(* IEC 61131-3 sources: sis-interlock-demo/tests/POUs/Generated/FB_CemGen02_Test, 41 files *)

(* ---- FB_CemGen02_Test.decl.st ---- *)
// AUTO-GENERATED by cemgen 1.0.0 — не редактировать: правьте матрицу и запустите
//   python -m cemgen generate <файл матрицы .csv или .xlsx>
// Матрица: SIS-V101-CEM, объект V-101, ревизия B от 2026-10-19, SHA-256 сетки df2ed4841a9453ca
// Назначение: набор coUnit: сценарии по матрице SIS-V101-CEM, тесты 41–80 (DESIGN.md, 12.4).
//             Ожидаемые значения — эталонная модель cemgen. Стенд FB_SisHarness — по экземпляру на
//             тест.
// Автор:      kr0nsch; код — генератор cemgen
// Версия:     1.0.0
// Документ:   docs/DESIGN.md, раздел «10. Генератор cemgen»; docs/cause_effect_matrix.md
// ВНИМАНИЕ:   код демонстрационный и не предназначен для систем безопасности. Реальная ПАЗ требует
//             определения SIL, сертифицированных аппаратных и программных средств и валидации по
//             ГОСТ Р МЭК 61511.
FUNCTION_BLOCK FB_CemGen02_Test EXTENDS coUnit.FB_TestSuite
VAR
    fbH001 : FB_SisHarness;   // Matrix_ASHH104Override_Denied
    fbH002 : FB_SisHarness;   // Matrix_ASHH104Reset_OnlyAfterClear
    fbH003 : FB_SisHarness;   // Matrix_ASHH104ChannelInvalid_MatchesPolicy
    fbH004 : FB_SisHarness;   // Matrix_ASHH104Bypass_ExpiresBackToVoting
    fbH005 : FB_SisHarness;   // Matrix_BSH105Demand_TripsOwnEffects
    fbH006 : FB_SisHarness;   // Matrix_BSH105Override_Denied
    fbH007 : FB_SisHarness;   // Matrix_BSH105Reset_OnlyAfterClear
    fbH008 : FB_SisHarness;   // Matrix_BSH105ChannelInvalid_MatchesPolicy
    fbH009 : FB_SisHarness;   // Matrix_BSH105Bypass_ExpiresBackToVoting
    fbH010 : FB_SisHarness;   // Matrix_HS106Demand_TripsOwnEffects
    fbH011 : FB_SisHarness;   // Matrix_HS106Override_Denied
    fbH012 : FB_SisHarness;   // Matrix_HS106Reset_OnlyAfterClear
    fbH013 : FB_SisHarness;   // Matrix_HS106ChannelInvalid_MatchesPolicy
    fbH014 : FB_SisHarness;   // Matrix_HS106Bypass_Denied
    fbH015 : FB_SisHarness;   // Matrix_PSLL108Demand_TripsOwnEffects
    fbH016 : FB_SisHarness;   // Matrix_PSLL108Delay_TripsExactlyAtDelay
    fbH017 : FB_SisHarness;   // Matrix_PSLL108Override_ExpiresThenTrips
    fbH018 : FB_SisHarness;   // Matrix_PSLL108Override_ClearsAfterConfirm
    fbH019 : FB_SisHarness;   // Matrix_PSLL108Override_DemandBackRestartsConfirm
    fbH020 : FB_SisHarness;   // Matrix_PSLL108Override_ExpiryBoundsConfirm
    fbH021 : FB_SisHarness;   // Matrix_PSLL108Override_ClearedThenDelayTrips
    fbH022 : FB_SisHarness;   // Matrix_PSLL108Reset_OnlyAfterClear
    fbH023 : FB_SisHarness;   // Matrix_PSLL108ChannelInvalid_MatchesPolicy
    fbH024 : FB_SisHarness;   // Matrix_PSLL108Bypass_ExpiresBackToVoting
    fbH025 : FB_SisHarness;   // Matrix_ESL109Demand_TripsOwnEffects
    fbH026 : FB_SisHarness;   // Matrix_ESL109Delay_TripsExactlyAtDelay
    fbH027 : FB_SisHarness;   // Matrix_ESL109Override_Denied
    fbH028 : FB_SisHarness;   // Matrix_ESL109Reset_OnlyAfterClear
    fbH029 : FB_SisHarness;   // Matrix_ESL109ChannelInvalid_MatchesPolicy
    fbH030 : FB_SisHarness;   // Matrix_ESL109Bypass_Denied
    fbH031 : FB_SisHarness;   // Matrix_FirstOutPSHH101ThenPSLL101_RecordsFirst
    fbH032 : FB_SisHarness;   // Matrix_FirstOutPSLL101ThenLSHH102_RecordsFirst
    fbH033 : FB_SisHarness;   // Matrix_FirstOutLSHH102ThenLSLL102_RecordsFirst
    fbH034 : FB_SisHarness;   // Matrix_FirstOutLSLL102ThenTSHH103_RecordsFirst
    fbH035 : FB_SisHarness;   // Matrix_FirstOutTSHH103ThenASHH104_RecordsFirst
    fbH036 : FB_SisHarness;   // Matrix_FirstOutASHH104ThenBSH105_RecordsFirst
    fbH037 : FB_SisHarness;   // Matrix_FirstOutBSH105ThenHS106_RecordsFirst
    fbH038 : FB_SisHarness;   // Matrix_FirstOutHS106ThenPSLL108_RecordsFirst
    fbH039 : FB_SisHarness;   // Matrix_FirstOutPSLL108ThenESL109_RecordsFirst
    fbH040 : FB_SisHarness;   // Matrix_FirstOutESL109ThenPSHH101_RecordsFirst
END_VAR

(* ---- ASHH104BypassExpiresBackToVoting.method.decl.st ---- *)
// AUTO-GENERATED by cemgen 1.0.0 — не редактировать: правьте матрицу и запустите
//   python -m cemgen generate <файл матрицы .csv или .xlsx>
// Матрица: SIS-V101-CEM, объект V-101, ревизия B от 2026-10-19, SHA-256 сетки df2ed4841a9453ca
// Назначение: тест Matrix_ASHH104Bypass_ExpiresBackToVoting набора FB_CemGen02_Test (сценарий по
//             матрице, DESIGN.md, 12.4).
// Автор:      kr0nsch; код — генератор cemgen
// Версия:     1.0.0
// Документ:   docs/DESIGN.md, раздел «10. Генератор cemgen»; docs/cause_effect_matrix.md
// ВНИМАНИЕ:   код демонстрационный и не предназначен для систем безопасности. Реальная ПАЗ требует
//             определения SIL, сертифицированных аппаратных и программных средств и валидации по
//             ГОСТ Р МЭК 61511.
// Причина 6 ASHH104: ключ разрешения байпасов, байпас AT104A → Active; канал недостоверен → Bypassed,
// не сработало; на t0 + 8 ч − шаг — Active; ровно на t0 + 8 ч — Expired, BypassExpired, канал Invalid;
// далее — по эталонной модели.
METHOD PRIVATE ASHH104BypassExpiresBackToVoting
VAR
    xArmed : BOOL;           // стенд взведён: все следствия под напряжением после сброса
    stVs   : ST_VotingSts;   // копия состояния группы голосования
END_VAR

(* ---- ASHH104ChannelInvalidMatchesPolicy.method.decl.st ---- *)
// AUTO-GENERATED by cemgen 1.0.0 — не редактировать: правьте матрицу и запустите
//   python -m cemgen generate <файл матрицы .csv или .xlsx>
// Матрица: SIS-V101-CEM, объект V-101, ревизия B от 2026-10-19, SHA-256 сетки df2ed4841a9453ca
// Назначение: тест Matrix_ASHH104ChannelInvalid_MatchesPolicy набора FB_CemGen02_Test (сценарий по
//             матрице, DESIGN.md, 12.4).
// Автор:      kr0nsch; код — генератор cemgen
// Версия:     1.0.0
// Документ:   docs/DESIGN.md, раздел «10. Генератор cemgen»; docs/cause_effect_matrix.md
// ВНИМАНИЕ:   код демонстрационный и не предназначен для систем безопасности. Реальная ПАЗ требует
//             определения SIL, сертифицированных аппаратных и программных средств и валидации по
//             ГОСТ Р МЭК 61511.
// Причина 6 ASHH104 (2oo3, DegradeSafe): канал AT104A недостоверен → действующая схема и срабатывание
// по политике деградации; если не сработало — требование на AT104B → по эталонной модели.
METHOD PRIVATE ASHH104ChannelInvalidMatchesPolicy
VAR
    xArmed : BOOL;           // стенд взведён: все следствия под напряжением после сброса
    stVs   : ST_VotingSts;   // копия состояния группы голосования
END_VAR

(* ---- ASHH104OverrideDenied.method.decl.st ---- *)
// AUTO-GENERATED by cemgen 1.0.0 — не редактировать: правьте матрицу и запустите
//   python -m cemgen generate <файл матрицы .csv или .xlsx>
// Матрица: SIS-V101-CEM, объект V-101, ревизия B от 2026-10-19, SHA-256 сетки df2ed4841a9453ca
// Назначение: тест Matrix_ASHH104Override_Denied набора FB_CemGen02_Test (сценарий по матрице,
//             DESIGN.md, 12.4).
// Автор:      kr0nsch; код — генератор cemgen
// Версия:     1.0.0
// Документ:   docs/DESIGN.md, раздел «10. Генератор cemgen»; docs/cause_effect_matrix.md
// ВНИМАНИЕ:   код демонстрационный и не предназначен для систем безопасности. Реальная ПАЗ требует
//             определения SIL, сертифицированных аппаратных и программных средств и валидации по
//             ГОСТ Р МЭК 61511.
// Причина 6 ASHH104 без разрешённого обхода: ключ разрешения обходов, запрос → последнее событие
// OverrideDenied, обхода нет; требование → срабатывание после задержки.
METHOD PRIVATE ASHH104OverrideDenied
VAR
    xArmed : BOOL;          // стенд взведён: все следствия под напряжением после сброса
    stEv   : ST_SisEvent;   // последнее событие журнала
END_VAR

(* ---- ASHH104ResetOnlyAfterClear.method.decl.st ---- *)
// AUTO-GENERATED by cemgen 1.0.0 — не редактировать: правьте матрицу и запустите
//   python -m cemgen generate <файл матрицы .csv или .xlsx>
// Матрица: SIS-V101-CEM, объект V-101, ревизия B от 2026-10-19, SHA-256 сетки df2ed4841a9453ca
// Назначение: тест Matrix_ASHH104Reset_OnlyAfterClear набора FB_CemGen02_Test (сценарий по матрице,
//             DESIGN.md, 12.4).
// Автор:      kr0nsch; код — генератор cemgen
// Версия:     1.0.0
// Документ:   docs/DESIGN.md, раздел «10. Генератор cemgen»; docs/cause_effect_matrix.md
// ВНИМАНИЕ:   код демонстрационный и не предназначен для систем безопасности. Реальная ПАЗ требует
//             определения SIL, сертифицированных аппаратных и программных средств и валидации по
//             ГОСТ Р МЭК 61511.
// Причина 6 ASHH104: срабатывание; сброс при требовании → ResetDenied, блокирует ASHH104, следствия
// обесточены; норма → следствия всё ещё обесточены (фиксация); сброс → все следствия под напряжением.
METHOD PRIVATE ASHH104ResetOnlyAfterClear
VAR
    xArmed : BOOL;          // стенд взведён: все следствия под напряжением после сброса
    stEv   : ST_SisEvent;   // последнее событие журнала
END_VAR

(* ---- BSH105BypassExpiresBackToVoting.method.decl.st ---- *)
// AUTO-GENERATED by cemgen 1.0.0 — не редактировать: правьте матрицу и запустите
//   python -m cemgen generate <файл матрицы .csv или .xlsx>
// Матрица: SIS-V101-CEM, объект V-101, ревизия B от 2026-10-19, SHA-256 сетки df2ed4841a9453ca
// Назначение: тест Matrix_BSH105Bypass_ExpiresBackToVoting набора FB_CemGen02_Test (сценарий по
//             матрице, DESIGN.md, 12.4).
// Автор:      kr0nsch; код — генератор cemgen
// Версия:     1.0.0
// Документ:   docs/DESIGN.md, раздел «10. Генератор cemgen»; docs/cause_effect_matrix.md
// ВНИМАНИЕ:   код демонстрационный и не предназначен для систем безопасности. Реальная ПАЗ требует
//             определения SIL, сертифицированных аппаратных и программных средств и валидации по
//             ГОСТ Р МЭК 61511.
// Причина 7 BSH105: ключ разрешения байпасов, байпас BS105A → Active; канал недостоверен → Bypassed,
// не сработало; на t0 + 8 ч − шаг — Active; ровно на t0 + 8 ч — Expired, BypassExpired, канал Invalid;
// далее — по эталонной модели.
METHOD PRIVATE BSH105BypassExpiresBackToVoting
VAR
    xArmed : BOOL;           // стенд взведён: все следствия под напряжением после сброса
    stVs   : ST_VotingSts;   // копия состояния группы голосования
END_VAR

(* ---- BSH105ChannelInvalidMatchesPolicy.method.decl.st ---- *)
// AUTO-GENERATED by cemgen 1.0.0 — не редактировать: правьте матрицу и запустите
//   python -m cemgen generate <файл матрицы .csv или .xlsx>
// Матрица: SIS-V101-CEM, объект V-101, ревизия B от 2026-10-19, SHA-256 сетки df2ed4841a9453ca
// Назначение: тест Matrix_BSH105ChannelInvalid_MatchesPolicy набора FB_CemGen02_Test (сценарий по
//             матрице, DESIGN.md, 12.4).
// Автор:      kr0nsch; код — генератор cemgen
// Версия:     1.0.0
// Документ:   docs/DESIGN.md, раздел «10. Генератор cemgen»; docs/cause_effect_matrix.md
// ВНИМАНИЕ:   код демонстрационный и не предназначен для систем безопасности. Реальная ПАЗ требует
//             определения SIL, сертифицированных аппаратных и программных средств и валидации по
//             ГОСТ Р МЭК 61511.
// Причина 7 BSH105 (1oo2, DegradeSafe): канал BS105A недостоверен → действующая схема и срабатывание
// по политике деградации; если не сработало — требование на BS105B → по эталонной модели.
METHOD PRIVATE BSH105ChannelInvalidMatchesPolicy
VAR
    xArmed : BOOL;           // стенд взведён: все следствия под напряжением после сброса
    stVs   : ST_VotingSts;   // копия состояния группы голосования
END_VAR

(* ---- BSH105DemandTripsOwnEffects.method.decl.st ---- *)
// AUTO-GENERATED by cemgen 1.0.0 — не редактировать: правьте матрицу и запустите
//   python -m cemgen generate <файл матрицы .csv или .xlsx>
// Матрица: SIS-V101-CEM, объект V-101, ревизия B от 2026-10-19, SHA-256 сетки df2ed4841a9453ca
// Назначение: тест Matrix_BSH105Demand_TripsOwnEffects набора FB_CemGen02_Test (сценарий по
//             матрице, DESIGN.md, 12.4).
// Автор:      kr0nsch; код — генератор cemgen
// Версия:     1.0.0
// Документ:   docs/DESIGN.md, раздел «10. Генератор cemgen»; docs/cause_effect_matrix.md
// ВНИМАНИЕ:   код демонстрационный и не предназначен для систем безопасности. Реальная ПАЗ требует
//             определения SIL, сертифицированных аппаратных и программных средств и валидации по
//             ГОСТ Р МЭК 61511.
// Причина 7 BSH105 (1oo2, задержка 0 с): требование BS105A, BS105B = 0 отключает ESDV101, BDV101,
// ESDV102, P101A, P101B, H101, UA110; остальные следствия под напряжением; первопричина BSH105.
METHOD PRIVATE BSH105DemandTripsOwnEffects
VAR
    xArmed : BOOL;   // стенд взведён: все следствия под напряжением после сброса
END_VAR

(* ---- BSH105OverrideDenied.method.decl.st ---- *)
// AUTO-GENERATED by cemgen 1.0.0 — не редактировать: правьте матрицу и запустите
//   python -m cemgen generate <файл матрицы .csv или .xlsx>
// Матрица: SIS-V101-CEM, объект V-101, ревизия B от 2026-10-19, SHA-256 сетки df2ed4841a9453ca
// Назначение: тест Matrix_BSH105Override_Denied набора FB_CemGen02_Test (сценарий по матрице,
//             DESIGN.md, 12.4).
// Автор:      kr0nsch; код — генератор cemgen
// Версия:     1.0.0
// Документ:   docs/DESIGN.md, раздел «10. Генератор cemgen»; docs/cause_effect_matrix.md
// ВНИМАНИЕ:   код демонстрационный и не предназначен для систем безопасности. Реальная ПАЗ требует
//             определения SIL, сертифицированных аппаратных и программных средств и валидации по
//             ГОСТ Р МЭК 61511.
// Причина 7 BSH105 без разрешённого обхода: ключ разрешения обходов, запрос → последнее событие
// OverrideDenied, обхода нет; требование → срабатывание после задержки.
METHOD PRIVATE BSH105OverrideDenied
VAR
    xArmed : BOOL;          // стенд взведён: все следствия под напряжением после сброса
    stEv   : ST_SisEvent;   // последнее событие журнала
END_VAR

(* ---- BSH105ResetOnlyAfterClear.method.decl.st ---- *)
// AUTO-GENERATED by cemgen 1.0.0 — не редактировать: правьте матрицу и запустите
//   python -m cemgen generate <файл матрицы .csv или .xlsx>
// Матрица: SIS-V101-CEM, объект V-101, ревизия B от 2026-10-19, SHA-256 сетки df2ed4841a9453ca
// Назначение: тест Matrix_BSH105Reset_OnlyAfterClear набора FB_CemGen02_Test (сценарий по матрице,
//             DESIGN.md, 12.4).
// Автор:      kr0nsch; код — генератор cemgen
// Версия:     1.0.0
// Документ:   docs/DESIGN.md, раздел «10. Генератор cemgen»; docs/cause_effect_matrix.md
// ВНИМАНИЕ:   код демонстрационный и не предназначен для систем безопасности. Реальная ПАЗ требует
//             определения SIL, сертифицированных аппаратных и программных средств и валидации по
//             ГОСТ Р МЭК 61511.
// Причина 7 BSH105: срабатывание; сброс при требовании → ResetDenied, блокирует BSH105, следствия
// обесточены; норма → следствия всё ещё обесточены (фиксация); сброс → все следствия под напряжением.
METHOD PRIVATE BSH105ResetOnlyAfterClear
VAR
    xArmed : BOOL;          // стенд взведён: все следствия под напряжением после сброса
    stEv   : ST_SisEvent;   // последнее событие журнала
END_VAR

(* ---- ESL109BypassDenied.method.decl.st ---- *)
// AUTO-GENERATED by cemgen 1.0.0 — не редактировать: правьте матрицу и запустите
//   python -m cemgen generate <файл матрицы .csv или .xlsx>
// Матрица: SIS-V101-CEM, объект V-101, ревизия B от 2026-10-19, SHA-256 сетки df2ed4841a9453ca
// Назначение: тест Matrix_ESL109Bypass_Denied набора FB_CemGen02_Test (сценарий по матрице,
//             DESIGN.md, 12.4).
// Автор:      kr0nsch; код — генератор cemgen
// Версия:     1.0.0
// Документ:   docs/DESIGN.md, раздел «10. Генератор cemgen»; docs/cause_effect_matrix.md
// ВНИМАНИЕ:   код демонстрационный и не предназначен для систем безопасности. Реальная ПАЗ требует
//             определения SIL, сертифицированных аппаратных и программных средств и валидации по
//             ГОСТ Р МЭК 61511.
// Причина 10 ESL109: байпас запрещён (bypass_max = 0); ключ разрешения байпасов, запрос байпаса ES109
// → Denied, событие BypassDenied с номером канала.
METHOD PRIVATE ESL109BypassDenied
VAR
    xArmed : BOOL;           // стенд взведён: все следствия под напряжением после сброса
    stVs   : ST_VotingSts;   // копия состояния группы голосования
    stEv   : ST_SisEvent;    // последнее событие журнала
END_VAR

(* ---- ESL109ChannelInvalidMatchesPolicy.method.decl.st ---- *)
// AUTO-GENERATED by cemgen 1.0.0 — не редактировать: правьте матрицу и запустите
//   python -m cemgen generate <файл матрицы .csv или .xlsx>
// Матрица: SIS-V101-CEM, объект V-101, ревизия B от 2026-10-19, SHA-256 сетки df2ed4841a9453ca
// Назначение: тест Matrix_ESL109ChannelInvalid_MatchesPolicy набора FB_CemGen02_Test (сценарий по
//             матрице, DESIGN.md, 12.4).
// Автор:      kr0nsch; код — генератор cemgen
// Версия:     1.0.0
// Документ:   docs/DESIGN.md, раздел «10. Генератор cemgen»; docs/cause_effect_matrix.md
// ВНИМАНИЕ:   код демонстрационный и не предназначен для систем безопасности. Реальная ПАЗ требует
//             определения SIL, сертифицированных аппаратных и программных средств и валидации по
//             ГОСТ Р МЭК 61511.
// Причина 10 ESL109 (1oo1, VoteTrip): канал ES109 недостоверен → действующая схема и срабатывание по
// политике деградации; если не сработало — требование на втором канале → по эталонной модели.
METHOD PRIVATE ESL109ChannelInvalidMatchesPolicy
VAR
    xArmed : BOOL;           // стенд взведён: все следствия под напряжением после сброса
    stVs   : ST_VotingSts;   // копия состояния группы голосования
END_VAR

(* ---- ESL109DelayTripsExactlyAtDelay.method.decl.st ---- *)
// AUTO-GENERATED by cemgen 1.0.0 — не редактировать: правьте матрицу и запустите
//   python -m cemgen generate <файл матрицы .csv или .xlsx>
// Матрица: SIS-V101-CEM, объект V-101, ревизия B от 2026-10-19, SHA-256 сетки df2ed4841a9453ca
// Назначение: тест Matrix_ESL109Delay_TripsExactlyAtDelay набора FB_CemGen02_Test (сценарий по
//             матрице, DESIGN.md, 12.4).
// Автор:      kr0nsch; код — генератор cemgen
// Версия:     1.0.0
// Документ:   docs/DESIGN.md, раздел «10. Генератор cemgen»; docs/cause_effect_matrix.md
// ВНИМАНИЕ:   код демонстрационный и не предназначен для систем безопасности. Реальная ПАЗ требует
//             определения SIL, сертифицированных аппаратных и программных средств и валидации по
//             ГОСТ Р МЭК 61511.
// Причина 10 ESL109: требование в t0; на t0 + 2 с − шаг не зафиксирована, следствия под напряжением;
// ровно на t0 + 2 с — зафиксирована, ltFirstOut = t0 + задержка.
METHOD PRIVATE ESL109DelayTripsExactlyAtDelay
VAR
    xArmed : BOOL;    // стенд взведён: все следствия под напряжением после сброса
    ltT0   : LTIME;   // момент t0 по подменному времени стенда
END_VAR

(* ---- ESL109DemandTripsOwnEffects.method.decl.st ---- *)
// AUTO-GENERATED by cemgen 1.0.0 — не редактировать: правьте матрицу и запустите
//   python -m cemgen generate <файл матрицы .csv или .xlsx>
// Матрица: SIS-V101-CEM, объект V-101, ревизия B от 2026-10-19, SHA-256 сетки df2ed4841a9453ca
// Назначение: тест Matrix_ESL109Demand_TripsOwnEffects набора FB_CemGen02_Test (сценарий по
//             матрице, DESIGN.md, 12.4).
// Автор:      kr0nsch; код — генератор cemgen
// Версия:     1.0.0
// Документ:   docs/DESIGN.md, раздел «10. Генератор cemgen»; docs/cause_effect_matrix.md
// ВНИМАНИЕ:   код демонстрационный и не предназначен для систем безопасности. Реальная ПАЗ требует
//             определения SIL, сертифицированных аппаратных и программных средств и валидации по
//             ГОСТ Р МЭК 61511.
// Причина 10 ESL109 (1oo1, задержка 2 с): требование ES109 = 0 отключает P101A, P101B, H101, UA110;
// остальные следствия под напряжением; первопричина ESL109.
METHOD PRIVATE ESL109DemandTripsOwnEffects
VAR
    xArmed : BOOL;   // стенд взведён: все следствия под напряжением после сброса
END_VAR

(* ---- ESL109OverrideDenied.method.decl.st ---- *)
// AUTO-GENERATED by cemgen 1.0.0 — не редактировать: правьте матрицу и запустите
//   python -m cemgen generate <файл матрицы .csv или .xlsx>
// Матрица: SIS-V101-CEM, объект V-101, ревизия B от 2026-10-19, SHA-256 сетки df2ed4841a9453ca
// Назначение: тест Matrix_ESL109Override_Denied набора FB_CemGen02_Test (сценарий по матрице,
//             DESIGN.md, 12.4).
// Автор:      kr0nsch; код — генератор cemgen
// Версия:     1.0.0
// Документ:   docs/DESIGN.md, раздел «10. Генератор cemgen»; docs/cause_effect_matrix.md
// ВНИМАНИЕ:   код демонстрационный и не предназначен для систем безопасности. Реальная ПАЗ требует
//             определения SIL, сертифицированных аппаратных и программных средств и валидации по
//             ГОСТ Р МЭК 61511.
// Причина 10 ESL109 без разрешённого обхода: ключ разрешения обходов, запрос → последнее событие
// OverrideDenied, обхода нет; требование → срабатывание после задержки.
METHOD PRIVATE ESL109OverrideDenied
VAR
    xArmed : BOOL;          // стенд взведён: все следствия под напряжением после сброса
    stEv   : ST_SisEvent;   // последнее событие журнала
END_VAR

(* ---- ESL109ResetOnlyAfterClear.method.decl.st ---- *)
// AUTO-GENERATED by cemgen 1.0.0 — не редактировать: правьте матрицу и запустите
//   python -m cemgen generate <файл матрицы .csv или .xlsx>
// Матрица: SIS-V101-CEM, объект V-101, ревизия B от 2026-10-19, SHA-256 сетки df2ed4841a9453ca
// Назначение: тест Matrix_ESL109Reset_OnlyAfterClear набора FB_CemGen02_Test (сценарий по матрице,
//             DESIGN.md, 12.4).
// Автор:      kr0nsch; код — генератор cemgen
// Версия:     1.0.0
// Документ:   docs/DESIGN.md, раздел «10. Генератор cemgen»; docs/cause_effect_matrix.md
// ВНИМАНИЕ:   код демонстрационный и не предназначен для систем безопасности. Реальная ПАЗ требует
//             определения SIL, сертифицированных аппаратных и программных средств и валидации по
//             ГОСТ Р МЭК 61511.
// Причина 10 ESL109: срабатывание; сброс при требовании → ResetDenied, блокирует ESL109, следствия
// обесточены; норма → следствия всё ещё обесточены (фиксация); сброс → все следствия под напряжением.
METHOD PRIVATE ESL109ResetOnlyAfterClear
VAR
    xArmed : BOOL;          // стенд взведён: все следствия под напряжением после сброса
    stEv   : ST_SisEvent;   // последнее событие журнала
END_VAR

(* ---- FirstOutASHH104ThenBSH105RecordsFirst.method.decl.st ---- *)
// AUTO-GENERATED by cemgen 1.0.0 — не редактировать: правьте матрицу и запустите
//   python -m cemgen generate <файл матрицы .csv или .xlsx>
// Матрица: SIS-V101-CEM, объект V-101, ревизия B от 2026-10-19, SHA-256 сетки df2ed4841a9453ca
// Назначение: тест Matrix_FirstOutASHH104ThenBSH105_RecordsFirst набора FB_CemGen02_Test (сценарий
//             по матрице, DESIGN.md, 12.4).
// Автор:      kr0nsch; код — генератор cemgen
// Версия:     1.0.0
// Документ:   docs/DESIGN.md, раздел «10. Генератор cemgen»; docs/cause_effect_matrix.md
// ВНИМАНИЕ:   код демонстрационный и не предназначен для систем безопасности. Реальная ПАЗ требует
//             определения SIL, сертифицированных аппаратных и программных средств и валидации по
//             ГОСТ Р МЭК 61511.
// Первопричина: требование ASHH104, фиксация через 2 с; затем требование BSH105, фиксация через 0 с →
// первопричина ASHH104, в маске первопричины только ASHH104, ltFirstOut — момент фиксации ASHH104,
// BSH105 — среди зафиксированных.
METHOD PRIVATE FirstOutASHH104ThenBSH105RecordsFirst
VAR
    xArmed : BOOL;    // стенд взведён: все следствия под напряжением после сброса
    ltT0   : LTIME;   // момент t0 по подменному времени стенда
END_VAR

(* ---- FirstOutBSH105ThenHS106RecordsFirst.method.decl.st ---- *)
// AUTO-GENERATED by cemgen 1.0.0 — не редактировать: правьте матрицу и запустите
//   python -m cemgen generate <файл матрицы .csv или .xlsx>
// Матрица: SIS-V101-CEM, объект V-101, ревизия B от 2026-10-19, SHA-256 сетки df2ed4841a9453ca
// Назначение: тест Matrix_FirstOutBSH105ThenHS106_RecordsFirst набора FB_CemGen02_Test (сценарий по
//             матрице, DESIGN.md, 12.4).
// Автор:      kr0nsch; код — генератор cemgen
// Версия:     1.0.0
// Документ:   docs/DESIGN.md, раздел «10. Генератор cemgen»; docs/cause_effect_matrix.md
// ВНИМАНИЕ:   код демонстрационный и не предназначен для систем безопасности. Реальная ПАЗ требует
//             определения SIL, сертифицированных аппаратных и программных средств и валидации по
//             ГОСТ Р МЭК 61511.
// Первопричина: требование BSH105, фиксация через 0 с; затем требование HS106, фиксация через 0 с →
// первопричина BSH105, в маске первопричины только BSH105, ltFirstOut — момент фиксации BSH105, HS106
// — среди зафиксированных.
METHOD PRIVATE FirstOutBSH105ThenHS106RecordsFirst
VAR
    xArmed : BOOL;    // стенд взведён: все следствия под напряжением после сброса
    ltT0   : LTIME;   // момент t0 по подменному времени стенда
END_VAR

(* ---- FirstOutESL109ThenPSHH101RecordsFirst.method.decl.st ---- *)
// AUTO-GENERATED by cemgen 1.0.0 — не редактировать: правьте матрицу и запустите
//   python -m cemgen generate <файл матрицы .csv или .xlsx>
// Матрица: SIS-V101-CEM, объект V-101, ревизия B от 2026-10-19, SHA-256 сетки df2ed4841a9453ca
// Назначение: тест Matrix_FirstOutESL109ThenPSHH101_RecordsFirst набора FB_CemGen02_Test (сценарий
//             по матрице, DESIGN.md, 12.4).
// Автор:      kr0nsch; код — генератор cemgen
// Версия:     1.0.0
// Документ:   docs/DESIGN.md, раздел «10. Генератор cemgen»; docs/cause_effect_matrix.md
// ВНИМАНИЕ:   код демонстрационный и не предназначен для систем безопасности. Реальная ПАЗ требует
//             определения SIL, сертифицированных аппаратных и программных средств и валидации по
//             ГОСТ Р МЭК 61511.
// Первопричина: требование ESL109, фиксация через 2 с; затем требование PSHH101, фиксация через 2 с →
// первопричина ESL109, в маске первопричины только ESL109, ltFirstOut — момент фиксации ESL109,
// PSHH101 — среди зафиксированных.
METHOD PRIVATE FirstOutESL109ThenPSHH101RecordsFirst
VAR
    xArmed : BOOL;    // стенд взведён: все следствия под напряжением после сброса
    ltT0   : LTIME;   // момент t0 по подменному времени стенда
END_VAR

(* ---- FirstOutHS106ThenPSLL108RecordsFirst.method.decl.st ---- *)
// AUTO-GENERATED by cemgen 1.0.0 — не редактировать: правьте матрицу и запустите
//   python -m cemgen generate <файл матрицы .csv или .xlsx>
// Матрица: SIS-V101-CEM, объект V-101, ревизия B от 2026-10-19, SHA-256 сетки df2ed4841a9453ca
// Назначение: тест Matrix_FirstOutHS106ThenPSLL108_RecordsFirst набора FB_CemGen02_Test (сценарий
//             по матрице, DESIGN.md, 12.4).
// Автор:      kr0nsch; код — генератор cemgen
// Версия:     1.0.0
// Документ:   docs/DESIGN.md, раздел «10. Генератор cemgen»; docs/cause_effect_matrix.md
// ВНИМАНИЕ:   код демонстрационный и не предназначен для систем безопасности. Реальная ПАЗ требует
//             определения SIL, сертифицированных аппаратных и программных средств и валидации по
//             ГОСТ Р МЭК 61511.
// Первопричина: требование HS106, фиксация через 0 с; затем требование PSLL108, фиксация через 10 с →
// первопричина HS106, в маске первопричины только HS106, ltFirstOut — момент фиксации HS106, PSLL108 —
// среди зафиксированных.
METHOD PRIVATE FirstOutHS106ThenPSLL108RecordsFirst
VAR
    xArmed : BOOL;    // стенд взведён: все следствия под напряжением после сброса
    ltT0   : LTIME;   // момент t0 по подменному времени стенда
END_VAR

(* ---- FirstOutLSHH102ThenLSLL102RecordsFirst.method.decl.st ---- *)
// AUTO-GENERATED by cemgen 1.0.0 — не редактировать: правьте матрицу и запустите
//   python -m cemgen generate <файл матрицы .csv или .xlsx>
// Матрица: SIS-V101-CEM, объект V-101, ревизия B от 2026-10-19, SHA-256 сетки df2ed4841a9453ca
// Назначение: тест Matrix_FirstOutLSHH102ThenLSLL102_RecordsFirst набора FB_CemGen02_Test (сценарий
//             по матрице, DESIGN.md, 12.4).
// Автор:      kr0nsch; код — генератор cemgen
// Версия:     1.0.0
// Документ:   docs/DESIGN.md, раздел «10. Генератор cemgen»; docs/cause_effect_matrix.md
// ВНИМАНИЕ:   код демонстрационный и не предназначен для систем безопасности. Реальная ПАЗ требует
//             определения SIL, сертифицированных аппаратных и программных средств и валидации по
//             ГОСТ Р МЭК 61511.
// Первопричина: требование LSHH102, фиксация через 3 с; затем требование LSLL102, фиксация через 5 с →
// первопричина LSHH102, в маске первопричины только LSHH102, ltFirstOut — момент фиксации LSHH102,
// LSLL102 — среди зафиксированных.
METHOD PRIVATE FirstOutLSHH102ThenLSLL102RecordsFirst
VAR
    xArmed : BOOL;    // стенд взведён: все следствия под напряжением после сброса
    ltT0   : LTIME;   // момент t0 по подменному времени стенда
END_VAR

(* ---- FirstOutLSLL102ThenTSHH103RecordsFirst.method.decl.st ---- *)
// AUTO-GENERATED by cemgen 1.0.0 — не редактировать: правьте матрицу и запустите
//   python -m cemgen generate <файл матрицы .csv или .xlsx>
// Матрица: SIS-V101-CEM, объект V-101, ревизия B от 2026-10-19, SHA-256 сетки df2ed4841a9453ca
// Назначение: тест Matrix_FirstOutLSLL102ThenTSHH103_RecordsFirst набора FB_CemGen02_Test (сценарий
//             по матрице, DESIGN.md, 12.4).
// Автор:      kr0nsch; код — генератор cemgen
// Версия:     1.0.0
// Документ:   docs/DESIGN.md, раздел «10. Генератор cemgen»; docs/cause_effect_matrix.md
// ВНИМАНИЕ:   код демонстрационный и не предназначен для систем безопасности. Реальная ПАЗ требует
//             определения SIL, сертифицированных аппаратных и программных средств и валидации по
//             ГОСТ Р МЭК 61511.
// Первопричина: требование LSLL102, фиксация через 5 с; затем требование TSHH103, фиксация через 5 с →
// первопричина LSLL102, в маске первопричины только LSLL102, ltFirstOut — момент фиксации LSLL102,
// TSHH103 — среди зафиксированных.
METHOD PRIVATE FirstOutLSLL102ThenTSHH103RecordsFirst
VAR
    xArmed : BOOL;    // стенд взведён: все следствия под напряжением после сброса
    ltT0   : LTIME;   // момент t0 по подменному времени стенда
END_VAR

(* ---- FirstOutPSHH101ThenPSLL101RecordsFirst.method.decl.st ---- *)
// AUTO-GENERATED by cemgen 1.0.0 — не редактировать: правьте матрицу и запустите
//   python -m cemgen generate <файл матрицы .csv или .xlsx>
// Матрица: SIS-V101-CEM, объект V-101, ревизия B от 2026-10-19, SHA-256 сетки df2ed4841a9453ca
// Назначение: тест Matrix_FirstOutPSHH101ThenPSLL101_RecordsFirst набора FB_CemGen02_Test (сценарий
//             по матрице, DESIGN.md, 12.4).
// Автор:      kr0nsch; код — генератор cemgen
// Версия:     1.0.0
// Документ:   docs/DESIGN.md, раздел «10. Генератор cemgen»; docs/cause_effect_matrix.md
// ВНИМАНИЕ:   код демонстрационный и не предназначен для систем безопасности. Реальная ПАЗ требует
//             определения SIL, сертифицированных аппаратных и программных средств и валидации по
//             ГОСТ Р МЭК 61511.
// Первопричина: требование PSHH101, фиксация через 2 с; затем требование PSLL101, фиксация через 5 с →
// первопричина PSHH101, в маске первопричины только PSHH101, ltFirstOut — момент фиксации PSHH101,
// PSLL101 — среди зафиксированных.
METHOD PRIVATE FirstOutPSHH101ThenPSLL101RecordsFirst
VAR
    xArmed : BOOL;    // стенд взведён: все следствия под напряжением после сброса
    ltT0   : LTIME;   // момент t0 по подменному времени стенда
END_VAR

(* ---- FirstOutPSLL101ThenLSHH102RecordsFirst.method.decl.st ---- *)
// AUTO-GENERATED by cemgen 1.0.0 — не редактировать: правьте матрицу и запустите
//   python -m cemgen generate <файл матрицы .csv или .xlsx>
// Матрица: SIS-V101-CEM, объект V-101, ревизия B от 2026-10-19, SHA-256 сетки df2ed4841a9453ca
// Назначение: тест Matrix_FirstOutPSLL101ThenLSHH102_RecordsFirst набора FB_CemGen02_Test (сценарий
//             по матрице, DESIGN.md, 12.4).
// Автор:      kr0nsch; код — генератор cemgen
// Версия:     1.0.0
// Документ:   docs/DESIGN.md, раздел «10. Генератор cemgen»; docs/cause_effect_matrix.md
// ВНИМАНИЕ:   код демонстрационный и не предназначен для систем безопасности. Реальная ПАЗ требует
//             определения SIL, сертифицированных аппаратных и программных средств и валидации по
//             ГОСТ Р МЭК 61511.
// Первопричина: требование PSLL101, фиксация через 5 с; затем требование LSHH102, фиксация через 3 с →
// первопричина PSLL101, в маске первопричины только PSLL101, ltFirstOut — момент фиксации PSLL101,
// LSHH102 — среди зафиксированных.
METHOD PRIVATE FirstOutPSLL101ThenLSHH102RecordsFirst
VAR
    xArmed : BOOL;    // стенд взведён: все следствия под напряжением после сброса
    ltT0   : LTIME;   // момент t0 по подменному времени стенда
END_VAR

(* ---- FirstOutPSLL108ThenESL109RecordsFirst.method.decl.st ---- *)
// AUTO-GENERATED by cemgen 1.0.0 — не редактировать: правьте матрицу и запустите
//   python -m cemgen generate <файл матрицы .csv или .xlsx>
// Матрица: SIS-V101-CEM, объект V-101, ревизия B от 2026-10-19, SHA-256 сетки df2ed4841a9453ca
// Назначение: тест Matrix_FirstOutPSLL108ThenESL109_RecordsFirst набора FB_CemGen02_Test (сценарий
//             по матрице, DESIGN.md, 12.4).
// Автор:      kr0nsch; код — генератор cemgen
// Версия:     1.0.0
// Документ:   docs/DESIGN.md, раздел «10. Генератор cemgen»; docs/cause_effect_matrix.md
// ВНИМАНИЕ:   код демонстрационный и не предназначен для систем безопасности. Реальная ПАЗ требует
//             определения SIL, сертифицированных аппаратных и программных средств и валидации по
//             ГОСТ Р МЭК 61511.
// Первопричина: требование PSLL108, фиксация через 10 с; затем требование ESL109, фиксация через 2 с →
// первопричина PSLL108, в маске первопричины только PSLL108, ltFirstOut — момент фиксации PSLL108,
// ESL109 — среди зафиксированных.
METHOD PRIVATE FirstOutPSLL108ThenESL109RecordsFirst
VAR
    xArmed : BOOL;    // стенд взведён: все следствия под напряжением после сброса
    ltT0   : LTIME;   // момент t0 по подменному времени стенда
END_VAR

(* ---- FirstOutTSHH103ThenASHH104RecordsFirst.method.decl.st ---- *)
// AUTO-GENERATED by cemgen 1.0.0 — не редактировать: правьте матрицу и запустите
//   python -m cemgen generate <файл матрицы .csv или .xlsx>
// Матрица: SIS-V101-CEM, объект V-101, ревизия B от 2026-10-19, SHA-256 сетки df2ed4841a9453ca
// Назначение: тест Matrix_FirstOutTSHH103ThenASHH104_RecordsFirst набора FB_CemGen02_Test (сценарий
//             по матрице, DESIGN.md, 12.4).
// Автор:      kr0nsch; код — генератор cemgen
// Версия:     1.0.0
// Документ:   docs/DESIGN.md, раздел «10. Генератор cemgen»; docs/cause_effect_matrix.md
// ВНИМАНИЕ:   код демонстрационный и не предназначен для систем безопасности. Реальная ПАЗ требует
//             определения SIL, сертифицированных аппаратных и программных средств и валидации по
//             ГОСТ Р МЭК 61511.
// Первопричина: требование TSHH103, фиксация через 5 с; затем требование ASHH104, фиксация через 2 с →
// первопричина TSHH103, в маске первопричины только TSHH103, ltFirstOut — момент фиксации TSHH103,
// ASHH104 — среди зафиксированных.
METHOD PRIVATE FirstOutTSHH103ThenASHH104RecordsFirst
VAR
    xArmed : BOOL;    // стенд взведён: все следствия под напряжением после сброса
    ltT0   : LTIME;   // момент t0 по подменному времени стенда
END_VAR

(* ---- HS106BypassDenied.method.decl.st ---- *)
// AUTO-GENERATED by cemgen 1.0.0 — не редактировать: правьте матрицу и запустите
//   python -m cemgen generate <файл матрицы .csv или .xlsx>
// Матрица: SIS-V101-CEM, объект V-101, ревизия B от 2026-10-19, SHA-256 сетки df2ed4841a9453ca
// Назначение: тест Matrix_HS106Bypass_Denied набора FB_CemGen02_Test (сценарий по матрице,
//             DESIGN.md, 12.4).
// Автор:      kr0nsch; код — генератор cemgen
// Версия:     1.0.0
// Документ:   docs/DESIGN.md, раздел «10. Генератор cemgen»; docs/cause_effect_matrix.md
// ВНИМАНИЕ:   код демонстрационный и не предназначен для систем безопасности. Реальная ПАЗ требует
//             определения SIL, сертифицированных аппаратных и программных средств и валидации по
//             ГОСТ Р МЭК 61511.
// Причина 8 HS106: байпас запрещён (bypass_max = 0); ключ разрешения байпасов, запрос байпаса HS106A →
// Denied, событие BypassDenied с номером канала.
METHOD PRIVATE HS106BypassDenied
VAR
    xArmed : BOOL;           // стенд взведён: все следствия под напряжением после сброса
    stVs   : ST_VotingSts;   // копия состояния группы голосования
    stEv   : ST_SisEvent;    // последнее событие журнала
END_VAR

(* ---- HS106ChannelInvalidMatchesPolicy.method.decl.st ---- *)
// AUTO-GENERATED by cemgen 1.0.0 — не редактировать: правьте матрицу и запустите
//   python -m cemgen generate <файл матрицы .csv или .xlsx>
// Матрица: SIS-V101-CEM, объект V-101, ревизия B от 2026-10-19, SHA-256 сетки df2ed4841a9453ca
// Назначение: тест Matrix_HS106ChannelInvalid_MatchesPolicy набора FB_CemGen02_Test (сценарий по
//             матрице, DESIGN.md, 12.4).
// Автор:      kr0nsch; код — генератор cemgen
// Версия:     1.0.0
// Документ:   docs/DESIGN.md, раздел «10. Генератор cemgen»; docs/cause_effect_matrix.md
// ВНИМАНИЕ:   код демонстрационный и не предназначен для систем безопасности. Реальная ПАЗ требует
//             определения SIL, сертифицированных аппаратных и программных средств и валидации по
//             ГОСТ Р МЭК 61511.
// Причина 8 HS106 (1oo2, VoteTrip): канал HS106A недостоверен → действующая схема и срабатывание по
// политике деградации; если не сработало — требование на HS106B → по эталонной модели.
METHOD PRIVATE HS106ChannelInvalidMatchesPolicy
VAR
    xArmed : BOOL;           // стенд взведён: все следствия под напряжением после сброса
    stVs   : ST_VotingSts;   // копия состояния группы голосования
END_VAR

(* ---- HS106DemandTripsOwnEffects.method.decl.st ---- *)
// AUTO-GENERATED by cemgen 1.0.0 — не редактировать: правьте матрицу и запустите
//   python -m cemgen generate <файл матрицы .csv или .xlsx>
// Матрица: SIS-V101-CEM, объект V-101, ревизия B от 2026-10-19, SHA-256 сетки df2ed4841a9453ca
// Назначение: тест Matrix_HS106Demand_TripsOwnEffects набора FB_CemGen02_Test (сценарий по матрице,
//             DESIGN.md, 12.4).
// Автор:      kr0nsch; код — генератор cemgen
// Версия:     1.0.0
// Документ:   docs/DESIGN.md, раздел «10. Генератор cemgen»; docs/cause_effect_matrix.md
// ВНИМАНИЕ:   код демонстрационный и не предназначен для систем безопасности. Реальная ПАЗ требует
//             определения SIL, сертифицированных аппаратных и программных средств и валидации по
//             ГОСТ Р МЭК 61511.
// Причина 8 HS106 (1oo2, задержка 0 с): требование HS106A, HS106B = 0 отключает ESDV101, BDV101,
// ESDV102, P101A, P101B, H101, UA110; остальные следствия под напряжением; первопричина HS106.
METHOD PRIVATE HS106DemandTripsOwnEffects
VAR
    xArmed : BOOL;   // стенд взведён: все следствия под напряжением после сброса
END_VAR

(* ---- HS106OverrideDenied.method.decl.st ---- *)
// AUTO-GENERATED by cemgen 1.0.0 — не редактировать: правьте матрицу и запустите
//   python -m cemgen generate <файл матрицы .csv или .xlsx>
// Матрица: SIS-V101-CEM, объект V-101, ревизия B от 2026-10-19, SHA-256 сетки df2ed4841a9453ca
// Назначение: тест Matrix_HS106Override_Denied набора FB_CemGen02_Test (сценарий по матрице,
//             DESIGN.md, 12.4).
// Автор:      kr0nsch; код — генератор cemgen
// Версия:     1.0.0
// Документ:   docs/DESIGN.md, раздел «10. Генератор cemgen»; docs/cause_effect_matrix.md
// ВНИМАНИЕ:   код демонстрационный и не предназначен для систем безопасности. Реальная ПАЗ требует
//             определения SIL, сертифицированных аппаратных и программных средств и валидации по
//             ГОСТ Р МЭК 61511.
// Причина 8 HS106 без разрешённого обхода: ключ разрешения обходов, запрос → последнее событие
// OverrideDenied, обхода нет; требование → срабатывание после задержки.
METHOD PRIVATE HS106OverrideDenied
VAR
    xArmed : BOOL;          // стенд взведён: все следствия под напряжением после сброса
    stEv   : ST_SisEvent;   // последнее событие журнала
END_VAR

(* ---- HS106ResetOnlyAfterClear.method.decl.st ---- *)
// AUTO-GENERATED by cemgen 1.0.0 — не редактировать: правьте матрицу и запустите
//   python -m cemgen generate <файл матрицы .csv или .xlsx>
// Матрица: SIS-V101-CEM, объект V-101, ревизия B от 2026-10-19, SHA-256 сетки df2ed4841a9453ca
// Назначение: тест Matrix_HS106Reset_OnlyAfterClear набора FB_CemGen02_Test (сценарий по матрице,
//             DESIGN.md, 12.4).
// Автор:      kr0nsch; код — генератор cemgen
// Версия:     1.0.0
// Документ:   docs/DESIGN.md, раздел «10. Генератор cemgen»; docs/cause_effect_matrix.md
// ВНИМАНИЕ:   код демонстрационный и не предназначен для систем безопасности. Реальная ПАЗ требует
//             определения SIL, сертифицированных аппаратных и программных средств и валидации по
//             ГОСТ Р МЭК 61511.
// Причина 8 HS106: срабатывание; сброс при требовании → ResetDenied, блокирует HS106, следствия
// обесточены; норма → следствия всё ещё обесточены (фиксация); сброс → все следствия под напряжением.
METHOD PRIVATE HS106ResetOnlyAfterClear
VAR
    xArmed : BOOL;          // стенд взведён: все следствия под напряжением после сброса
    stEv   : ST_SisEvent;   // последнее событие журнала
END_VAR

(* ---- PSLL108BypassExpiresBackToVoting.method.decl.st ---- *)
// AUTO-GENERATED by cemgen 1.0.0 — не редактировать: правьте матрицу и запустите
//   python -m cemgen generate <файл матрицы .csv или .xlsx>
// Матрица: SIS-V101-CEM, объект V-101, ревизия B от 2026-10-19, SHA-256 сетки df2ed4841a9453ca
// Назначение: тест Matrix_PSLL108Bypass_ExpiresBackToVoting набора FB_CemGen02_Test (сценарий по
//             матрице, DESIGN.md, 12.4).
// Автор:      kr0nsch; код — генератор cemgen
// Версия:     1.0.0
// Документ:   docs/DESIGN.md, раздел «10. Генератор cemgen»; docs/cause_effect_matrix.md
// ВНИМАНИЕ:   код демонстрационный и не предназначен для систем безопасности. Реальная ПАЗ требует
//             определения SIL, сертифицированных аппаратных и программных средств и валидации по
//             ГОСТ Р МЭК 61511.
// Причина 9 PSLL108: ключ разрешения байпасов, байпас PS108A → Active; канал недостоверен → Bypassed,
// не сработало; на t0 + 4 ч − шаг — Active; ровно на t0 + 4 ч — Expired, BypassExpired, канал Invalid;
// далее — по эталонной модели.
METHOD PRIVATE PSLL108BypassExpiresBackToVoting
VAR
    xArmed : BOOL;           // стенд взведён: все следствия под напряжением после сброса
    stVs   : ST_VotingSts;   // копия состояния группы голосования
END_VAR

(* ---- PSLL108ChannelInvalidMatchesPolicy.method.decl.st ---- *)
// AUTO-GENERATED by cemgen 1.0.0 — не редактировать: правьте матрицу и запустите
//   python -m cemgen generate <файл матрицы .csv или .xlsx>
// Матрица: SIS-V101-CEM, объект V-101, ревизия B от 2026-10-19, SHA-256 сетки df2ed4841a9453ca
// Назначение: тест Matrix_PSLL108ChannelInvalid_MatchesPolicy набора FB_CemGen02_Test (сценарий по
//             матрице, DESIGN.md, 12.4).
// Автор:      kr0nsch; код — генератор cemgen
// Версия:     1.0.0
// Документ:   docs/DESIGN.md, раздел «10. Генератор cemgen»; docs/cause_effect_matrix.md
// ВНИМАНИЕ:   код демонстрационный и не предназначен для систем безопасности. Реальная ПАЗ требует
//             определения SIL, сертифицированных аппаратных и программных средств и валидации по
//             ГОСТ Р МЭК 61511.
// Причина 9 PSLL108 (2oo2, DegradeSafe): канал PS108A недостоверен → действующая схема и срабатывание
// по политике деградации; если не сработало — требование на PS108B → по эталонной модели.
METHOD PRIVATE PSLL108ChannelInvalidMatchesPolicy
VAR
    xArmed : BOOL;           // стенд взведён: все следствия под напряжением после сброса
    stVs   : ST_VotingSts;   // копия состояния группы голосования
END_VAR

(* ---- PSLL108DelayTripsExactlyAtDelay.method.decl.st ---- *)
// AUTO-GENERATED by cemgen 1.0.0 — не редактировать: правьте матрицу и запустите
//   python -m cemgen generate <файл матрицы .csv или .xlsx>
// Матрица: SIS-V101-CEM, объект V-101, ревизия B от 2026-10-19, SHA-256 сетки df2ed4841a9453ca
// Назначение: тест Matrix_PSLL108Delay_TripsExactlyAtDelay набора FB_CemGen02_Test (сценарий по
//             матрице, DESIGN.md, 12.4).
// Автор:      kr0nsch; код — генератор cemgen
// Версия:     1.0.0
// Документ:   docs/DESIGN.md, раздел «10. Генератор cemgen»; docs/cause_effect_matrix.md
// ВНИМАНИЕ:   код демонстрационный и не предназначен для систем безопасности. Реальная ПАЗ требует
//             определения SIL, сертифицированных аппаратных и программных средств и валидации по
//             ГОСТ Р МЭК 61511.
// Причина 9 PSLL108: требование в t0; на t0 + 10 с − шаг не зафиксирована, следствия под напряжением;
// ровно на t0 + 10 с — зафиксирована, ltFirstOut = t0 + задержка.
METHOD PRIVATE PSLL108DelayTripsExactlyAtDelay
VAR
    xArmed : BOOL;    // стенд взведён: все следствия под напряжением после сброса
    ltT0   : LTIME;   // момент t0 по подменному времени стенда
END_VAR

(* ---- PSLL108DemandTripsOwnEffects.method.decl.st ---- *)
// AUTO-GENERATED by cemgen 1.0.0 — не редактировать: правьте матрицу и запустите
//   python -m cemgen generate <файл матрицы .csv или .xlsx>
// Матрица: SIS-V101-CEM, объект V-101, ревизия B от 2026-10-19, SHA-256 сетки df2ed4841a9453ca
// Назначение: тест Matrix_PSLL108Demand_TripsOwnEffects набора FB_CemGen02_Test (сценарий по
//             матрице, DESIGN.md, 12.4).
// Автор:      kr0nsch; код — генератор cemgen
// Версия:     1.0.0
// Документ:   docs/DESIGN.md, раздел «10. Генератор cemgen»; docs/cause_effect_matrix.md
// ВНИМАНИЕ:   код демонстрационный и не предназначен для систем безопасности. Реальная ПАЗ требует
//             определения SIL, сертифицированных аппаратных и программных средств и валидации по
//             ГОСТ Р МЭК 61511.
// Причина 9 PSLL108 (2oo2, задержка 10 с): требование PS108A, PS108B = 0 отключает ESDV101, ESDV102,
// P101A, P101B, H101, UA110; остальные следствия под напряжением; первопричина PSLL108.
METHOD PRIVATE PSLL108DemandTripsOwnEffects
VAR
    xArmed : BOOL;   // стенд взведён: все следствия под напряжением после сброса
END_VAR

(* ---- PSLL108OverrideClearedThenDelayTrips.method.decl.st ---- *)
// AUTO-GENERATED by cemgen 1.0.0 — не редактировать: правьте матрицу и запустите
//   python -m cemgen generate <файл матрицы .csv или .xlsx>
// Матрица: SIS-V101-CEM, объект V-101, ревизия B от 2026-10-19, SHA-256 сетки df2ed4841a9453ca
// Назначение: тест Matrix_PSLL108Override_ClearedThenDelayTrips набора FB_CemGen02_Test (сценарий
//             по матрице, DESIGN.md, 12.4).
// Автор:      kr0nsch; код — генератор cemgen
// Версия:     1.0.0
// Документ:   docs/DESIGN.md, раздел «10. Генератор cemgen»; docs/cause_effect_matrix.md
// ВНИМАНИЕ:   код демонстрационный и не предназначен для систем безопасности. Реальная ПАЗ требует
//             определения SIL, сертифицированных аппаратных и программных средств и валидации по
//             ГОСТ Р МЭК 61511.
// Причина 9 PSLL108 с задержкой 10 с: пусковой обход и требование в t0; через 10 с причина активна под
// обходом, не зафиксирована; норма; через 30 с — OverrideCleared; требование в t2 — на t2 + 10 с − шаг
// не зафиксирована (задержка отсчитывается заново), на t2 + 10 с — зафиксирована, первопричина
// PSLL108.
METHOD PRIVATE PSLL108OverrideClearedThenDelayTrips
VAR
    xArmed : BOOL;    // стенд взведён: все следствия под напряжением после сброса
    ltT0   : LTIME;   // момент t2 по подменному времени стенда
END_VAR

(* ---- PSLL108OverrideClearsAfterConfirm.method.decl.st ---- *)
// AUTO-GENERATED by cemgen 1.0.0 — не редактировать: правьте матрицу и запустите
//   python -m cemgen generate <файл матрицы .csv или .xlsx>
// Матрица: SIS-V101-CEM, объект V-101, ревизия B от 2026-10-19, SHA-256 сетки df2ed4841a9453ca
// Назначение: тест Matrix_PSLL108Override_ClearsAfterConfirm набора FB_CemGen02_Test (сценарий по
//             матрице, DESIGN.md, 12.4).
// Автор:      kr0nsch; код — генератор cemgen
// Версия:     1.0.0
// Документ:   docs/DESIGN.md, раздел «10. Генератор cemgen»; docs/cause_effect_matrix.md
// ВНИМАНИЕ:   код демонстрационный и не предназначен для систем безопасности. Реальная ПАЗ требует
//             определения SIL, сертифицированных аппаратных и программных средств и валидации по
//             ГОСТ Р МЭК 61511.
// Причина 9 PSLL108: пусковой обход и требование в t0; норма с t1 = t0 + шаг; на t1 + 30 с − шаг обход
// действует; ровно на t1 + 30 с (подтверждение нормы) — OverrideCleared, обхода нет, причина не
// зафиксирована, следствия под напряжением (R-12).
METHOD PRIVATE PSLL108OverrideClearsAfterConfirm
VAR
    xArmed : BOOL;   // стенд взведён: все следствия под напряжением после сброса
END_VAR

(* ---- PSLL108OverrideDemandBackRestartsConfirm.method.decl.st ---- *)
// AUTO-GENERATED by cemgen 1.0.0 — не редактировать: правьте матрицу и запустите
//   python -m cemgen generate <файл матрицы .csv или .xlsx>
// Матрица: SIS-V101-CEM, объект V-101, ревизия B от 2026-10-19, SHA-256 сетки df2ed4841a9453ca
// Назначение: тест Matrix_PSLL108Override_DemandBackRestartsConfirm набора FB_CemGen02_Test
//             (сценарий по матрице, DESIGN.md, 12.4).
// Автор:      kr0nsch; код — генератор cemgen
// Версия:     1.0.0
// Документ:   docs/DESIGN.md, раздел «10. Генератор cemgen»; docs/cause_effect_matrix.md
// ВНИМАНИЕ:   код демонстрационный и не предназначен для систем безопасности. Реальная ПАЗ требует
//             определения SIL, сертифицированных аппаратных и программных средств и валидации по
//             ГОСТ Р МЭК 61511.
// Причина 9 PSLL108: пусковой обход и требование в t0; норма с t1; ровно на t1 + 30 с, когда обход
// снялся бы, требование снова — обход действует, подтверждение нормы сброшено; норма с t2; на t2 + 30
// с − шаг обход действует; на t2 + 30 с — OverrideCleared.
METHOD PRIVATE PSLL108OverrideDemandBackRestartsConfirm
VAR
    xArmed : BOOL;   // стенд взведён: все следствия под напряжением после сброса
END_VAR

(* ---- PSLL108OverrideExpiresThenTrips.method.decl.st ---- *)
// AUTO-GENERATED by cemgen 1.0.0 — не редактировать: правьте матрицу и запустите
//   python -m cemgen generate <файл матрицы .csv или .xlsx>
// Матрица: SIS-V101-CEM, объект V-101, ревизия B от 2026-10-19, SHA-256 сетки df2ed4841a9453ca
// Назначение: тест Matrix_PSLL108Override_ExpiresThenTrips набора FB_CemGen02_Test (сценарий по
//             матрице, DESIGN.md, 12.4).
// Автор:      kr0nsch; код — генератор cemgen
// Версия:     1.0.0
// Документ:   docs/DESIGN.md, раздел «10. Генератор cemgen»; docs/cause_effect_matrix.md
// ВНИМАНИЕ:   код демонстрационный и не предназначен для систем безопасности. Реальная ПАЗ требует
//             определения SIL, сертифицированных аппаратных и программных средств и валидации по
//             ГОСТ Р МЭК 61511.
// Причина 9 PSLL108: ключ разрешения обходов, запрос пускового обхода и требование в одном вызове t0;
// до t0 + 10 мин − шаг обход действует, причина не зафиксирована; ровно на t0 + 10 мин —
// OverrideExpired, фиксация, первопричина PSLL108.
METHOD PRIVATE PSLL108OverrideExpiresThenTrips
VAR
    xArmed : BOOL;   // стенд взведён: все следствия под напряжением после сброса
END_VAR

(* ---- PSLL108OverrideExpiryBoundsConfirm.method.decl.st ---- *)
// AUTO-GENERATED by cemgen 1.0.0 — не редактировать: правьте матрицу и запустите
//   python -m cemgen generate <файл матрицы .csv или .xlsx>
// Матрица: SIS-V101-CEM, объект V-101, ревизия B от 2026-10-19, SHA-256 сетки df2ed4841a9453ca
// Назначение: тест Matrix_PSLL108Override_ExpiryBoundsConfirm набора FB_CemGen02_Test (сценарий по
//             матрице, DESIGN.md, 12.4).
// Автор:      kr0nsch; код — генератор cemgen
// Версия:     1.0.0
// Документ:   docs/DESIGN.md, раздел «10. Генератор cemgen»; docs/cause_effect_matrix.md
// ВНИМАНИЕ:   код демонстрационный и не предназначен для систем безопасности. Реальная ПАЗ требует
//             определения SIL, сертифицированных аппаратных и программных средств и валидации по
//             ГОСТ Р МЭК 61511.
// Причина 9 PSLL108: пусковой обход и требование в t0; норма с t0 + 9 мин 30 с + шаг — подтверждение
// (30 с) закончилось бы после срока; на t0 + 10 мин − шаг обход действует; ровно на t0 + 10 мин —
// OverrideExpired (срок — верхняя граница), OverrideCleared нет, причина не зафиксирована (требования
// нет).
METHOD PRIVATE PSLL108OverrideExpiryBoundsConfirm
VAR
    xArmed : BOOL;   // стенд взведён: все следствия под напряжением после сброса
END_VAR

(* ---- PSLL108ResetOnlyAfterClear.method.decl.st ---- *)
// AUTO-GENERATED by cemgen 1.0.0 — не редактировать: правьте матрицу и запустите
//   python -m cemgen generate <файл матрицы .csv или .xlsx>
// Матрица: SIS-V101-CEM, объект V-101, ревизия B от 2026-10-19, SHA-256 сетки df2ed4841a9453ca
// Назначение: тест Matrix_PSLL108Reset_OnlyAfterClear набора FB_CemGen02_Test (сценарий по матрице,
//             DESIGN.md, 12.4).
// Автор:      kr0nsch; код — генератор cemgen
// Версия:     1.0.0
// Документ:   docs/DESIGN.md, раздел «10. Генератор cemgen»; docs/cause_effect_matrix.md
// ВНИМАНИЕ:   код демонстрационный и не предназначен для систем безопасности. Реальная ПАЗ требует
//             определения SIL, сертифицированных аппаратных и программных средств и валидации по
//             ГОСТ Р МЭК 61511.
// Причина 9 PSLL108: срабатывание; сброс при требовании → ResetDenied, блокирует PSLL108, следствия
// обесточены; норма → следствия всё ещё обесточены (фиксация); сброс → все следствия под напряжением.
METHOD PRIVATE PSLL108ResetOnlyAfterClear
VAR
    xArmed : BOOL;          // стенд взведён: все следствия под напряжением после сброса
    stEv   : ST_SisEvent;   // последнее событие журнала
END_VAR
